TYPE "DT_PARAM_ALL"
VERSION : 0.1
   STRUCT
      NOM_VAL_AND_CTRL : "DT_PAR_NOM_VAL_AND_CTRL";
      CTRL_2 : "DT_PAR_CTRL_2";
      DEVICES : "DT_PAR_DEVICES";
      SUBSYSTEM_MEAS_1 : "DT_PAR_SUBSYSTEM_MEAS_1";
      SUBSYSTEM_MEAS_2 : "DT_PAR_SUBSYSTEM_MEAS_2";
      SUBSYSTEM_MEAS_3 : "DT_PAR_SUBSYSTEM_MEAS_3";
      SUBSYSTEM_MEAS_4 : "DT_PAR_SUBSYSTEM_MEAS_4";
      SUB_SYSTEM_CTRL : "DT_PAR_SUB_SYSTEM_CTRL";
      SUB_SYSTEM_CTRL_2 : "DT_PAR_SUB_SYSTEM_CTRL_2";
      GEN_MEAS : "DT_PAR_GEN_MEAS";
      GEN_MEAS_2 : "DT_PAR_GEN_MEAS_2";
      GEN_SPEED : "DT_PAR_GEN_SPEED";
      GEN_WH_VIB : "DT_PAR_GEN_WH_VIB";
      GEN_EXC : "DT_PAR_GEN_EXC";
      TUR_POS_MEAS_1 : "DT_PAR_TUR_POS_MEAS_1";
      TUR_POS_MEAS_2 : "DT_PAR_TUR_POS_MEAS_2";
      TURBINE_1 : "DT_PAR_TURBINE_1";
      TURBINE_2 : "DT_PAR_TURBINE_2";
      TURBINE_3 : "DT_PAR_TURBINE_3";
      PID_WATER_LEVEL : "DT_PAR_PID_WATER_LEVEL";
      PID_WATER_PRESSURE : "DT_PAR_PID_WATER_PRESSURE";
      PID_ACTIVE_POWER : "DT_PAR_PID_ACTIVE_POWER";
      PID_SPEED : "DT_PAR_PID_SPEED";
      PID_FRANCIS_DISTRIBUTOR : "DT_PAR_PID_FRANCIS_DISTRIBUTOR";
      PID_KAPLAN_DISTRIBUTOR : "DT_PAR_PID_KAPLAN_DISTRIBUTOR";
      PID_KAPLAN_RUNNER : "DT_PAR_PID_KAPLAN_RUNNER";
      PID_CROSS_FLOW_VALVE_1 : "DT_PAR_PID_CROSS_FLOW_VALVE_1";
      PID_CROSS_FLOW_VALVE_2 : "DT_PAR_PID_CROSS_FLOW_VALVE_2";
      PID_PELTON_NOZZLE_1 : "DT_PAR_PID_PELTON_NOZZLE_1";
      PID_PELTON_NOZZLE_2 : "DT_PAR_PID_PELTON_NOZZLE_2";
      PID_PELTON_NOZZLE_3 : "DT_PAR_PID_PELTON_NOZZLE_3";
      PID_PELTON_NOZZLE_4 : "DT_PAR_PID_PELTON_NOZZLE_4";
      PID_PELTON_NOZZLE_5 : "DT_PAR_PID_PELTON_NOZZLE_5";
      PID_PELTON_NOZZLE_6 : "DT_PAR_PID_PELTON_NOZZLE_6";
      PID_PELTON_DEFLECTOR_1 : "DT_PAR_PID_PELTON_DEFLECTOR_1";
   END_STRUCT;

END_TYPE

